(* IEC 61131-3 sources: genai_codesys/tests/fixtures/codesys, 14 files *)

(* ---- custom_09_valid_declaration.st ---- *)
FUNCTION_BLOCK FB_JamMonitor
VAR_INPUT
    runCommand : BOOL;
    sensorPulse : BOOL;
    emergencyStop : BOOL;
    reset : BOOL;
END_VAR
VAR_OUTPUT
    motorRun : BOOL;
    jamAlarm : BOOL;
END_VAR
VAR
    watchdog : TON;
END_VAR

(* ---- fifo_fb_declaration.st ---- *)
FUNCTION_BLOCK FifoQueueProbe
VAR_IN_OUT
    item : DINT;
    buffer : ARRAY[1..10] OF DINT;
END_VAR
VAR_OUTPUT
    ok : BOOL;
END_VAR

(* ---- invalid_fb_declaration.st ---- *)
FUNCTION_BLOCK MotorControl
VAR_INPUT
    StartBtn : BOOL;
    StopBtn : BOOL;
    EStop : BOOL;
END_VAR
VAR_OUTPUT
    Motor : BOOL;
END_VAR

(* ---- public_18_valid_declaration.st ---- *)
FUNCTION_BLOCK FB_FIFOQueue
VAR_INPUT
    enqueue : BOOL;
    dequeue : BOOL;
    reset : BOOL;
END_VAR
VAR_OUTPUT
    elementCount : DINT;
    status : WORD;
END_VAR
VAR_IN_OUT
    item : DINT;
    buffer : ARRAY[1..10] OF DINT;
END_VAR
VAR
    head : DINT := 1;
    tail : DINT := 1;
    previousEnqueue : BOOL;
    previousDequeue : BOOL;
END_VAR

(* ---- special_fb_declaration.st ---- *)
FUNCTION_BLOCK PumpGroupControl
VAR_IN_OUT
    pumpGroup : ARRAY[1..5] OF ST_Pump;
END_VAR

(* ---- valid_fb_declaration.st ---- *)
FUNCTION_BLOCK MotorControl
VAR_INPUT
    StartBtn : BOOL;
    StopBtn : BOOL;
    EStop : BOOL;
END_VAR
VAR_OUTPUT
    Motor : BOOL;
END_VAR

(* ---- custom_09_valid_implementation.st ---- *)
IF reset AND NOT runCommand AND NOT emergencyStop THEN
    jamAlarm := FALSE;
END_IF;

motorRun := runCommand AND NOT emergencyStop AND NOT jamAlarm;
watchdog(IN := motorRun AND NOT sensorPulse, PT := T#2s);

IF watchdog.Q THEN
    jamAlarm := TRUE;
    motorRun := FALSE;
END_IF;

(* ---- invalid_declaration.st ---- *)
PROGRAM PLC_PRG
VAR
    StartBtn : BOOL;
    Motor : BOOL;
END_VAR

(* ---- invalid_fb_implementation.st ---- *)
IF StopBtn OR EStop THEN
    Motor := FALSE;
ELSIF StartBtn THEN
    Motor := MissingSignal;
END_IF;

(* ---- invalid_implementation.st ---- *)
IF StartBtn THEN
    Motor := TRUE
END_IF;

(* ---- public_18_valid_implementation.st ---- *)
IF reset THEN
    elementCount := 0;
    head := 1;
    tail := 1;
    status := 16#0000;
ELSIF enqueue AND NOT previousEnqueue THEN
    IF elementCount >= 10 THEN
        status := 16#8002;
    ELSE
        buffer[tail] := item;
        tail := tail + 1;
        IF tail > 10 THEN
            tail := 1;
        END_IF;
        elementCount := elementCount + 1;
        status := 16#0000;
    END_IF;
ELSIF dequeue AND NOT previousDequeue THEN
    IF elementCount <= 0 THEN
        status := 16#8001;
    ELSE
        item := buffer[head];
        head := head + 1;
        IF head > 10 THEN
            head := 1;
        END_IF;
        elementCount := elementCount - 1;
        status := 16#0000;
    END_IF;
END_IF;

previousEnqueue := enqueue;
previousDequeue := dequeue;

(* ---- valid_declaration.st ---- *)
PROGRAM PLC_PRG
VAR
    StartBtn : BOOL;
    StopBtn : BOOL;
    EStop : BOOL;
    Motor : BOOL;
END_VAR

(* ---- valid_fb_implementation.st ---- *)
IF StopBtn OR EStop THEN
    Motor := FALSE;
ELSIF StartBtn THEN
    Motor := TRUE;
END_IF;

(* ---- valid_implementation.st ---- *)
IF StopBtn OR EStop THEN
    Motor := FALSE;
ELSIF StartBtn THEN
    Motor := TRUE;
END_IF;
